FUNCTION_BLOCK FB_Valve IMPLEMENTS I_Valve
VAR_INPUT
	bClose	: BOOL;
END_VAR
VAR_OUTPUT
	bIsOpen	: BOOL;
END_VAR
VAR
	_eState	: E_ValveState;
	_nTicks	: UINT;
END_VAR

IF bClose THEN
	Act_Close();
END_IF
IF _eState = E_ValveState.Opening THEN
	_nTicks := _nTicks + 1;
	IF _nTicks >= 10 THEN
		_eState := E_ValveState.Open;
	END_IF
END_IF
bIsOpen := _eState = E_ValveState.Open;

METHOD Open : BOOL
VAR
END_VAR
IF _eState = E_ValveState.Closed THEN
	_eState := E_ValveState.Opening;
	_nTicks := 0;
END_IF
Open := _eState <> E_ValveState.Closed;
END_METHOD

PROPERTY State : E_ValveState
GET
State := _eState;
END_GET
SET
_eState := State;
END_SET
END_PROPERTY

ACTION Act_Close:
_eState := E_ValveState.Closed;
_nTicks := 0;
END_ACTION

END_FUNCTION_BLOCK

(* stored: Version 1.1.0.1, ProductVersion 3.1.4024.12
   POU FB_Valve: Id {90be5c88-da22-4202-bf6b-0788eb0769d5}, SpecialFunc None
   Folder Actions: Id {67d72acf-1e80-4c53-bb7f-868b743319fd}
   Method Open: Id {8e122aad-0321-4c46-a78b-aac38cef031a}
   Property State: Id {e68b2721-dac6-4526-9fac-83f157ff1574}
   Get Get: Id {f2de8de5-faaa-443f-bfa1-8deae8bbfea4}
   Set Set: Id {5031f7d9-b840-41b5-8b4e-e06696d82af7}
   Action Act_Close: Id {ae3481d1-5b24-42e6-86b7-8b071a0f8d86} *)
